FUNCTION_BLOCK SortingSafeSteps (* Standard safe-position sequence and its original timing. *)
  (* Standard: 61499-2 *)
  (* Version 3.0, 2026-11-12, sorting2n, sorting2n *)
  PACKAGE Main;
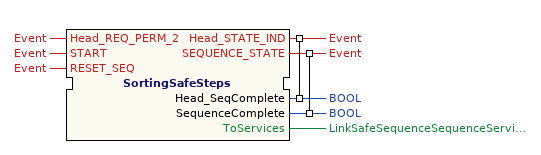
  EVENT_INPUT
    Head_REQ_PERM_2;
    START;
    RESET_SEQ;
  END_EVENT
  EVENT_OUTPUT
    Head_STATE_IND WITH Head_SeqComplete;
    SEQUENCE_STATE WITH SequenceComplete;
  END_EVENT
  VAR_OUTPUT
    Head_SeqComplete : BOOL;
    SequenceComplete : BOOL;
  END_VAR
  PLUGS
    ToServices : LinkSafeSequenceSequenceServices;
  END_PLUGS
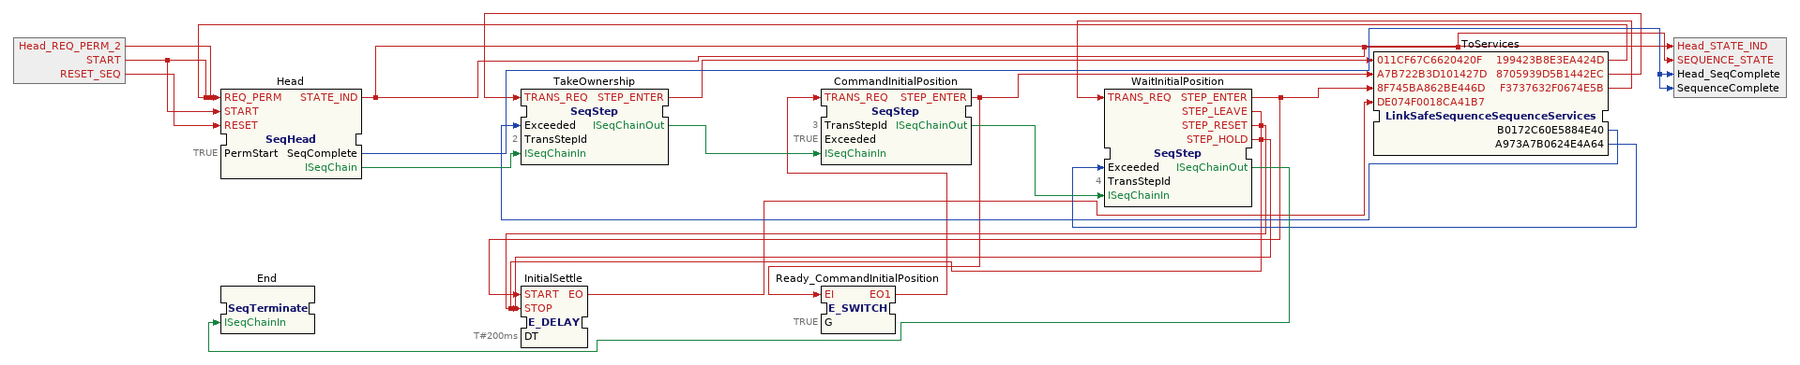
  FBS
    Head : SeqHead(PermStart := TRUE);
    End : SeqTerminate;
    TakeOwnership : SeqStep(TransStepId := 2);
    CommandInitialPosition : SeqStep(TransStepId := 3, Exceeded := TRUE);
    WaitInitialPosition : SeqStep(TransStepId := 4);
    InitialSettle : E_DELAY(DT := T#200ms);
    Ready_CommandInitialPosition : E_SWITCH(G := TRUE);
  END_FBS
  EVENT_CONNECTIONS
    Head.STATE_IND TO Head_STATE_IND;
    ToServices.199423B8E3EA424D TO Head.REQ_PERM;
    Head_REQ_PERM_2 TO Head.REQ_PERM;
    TakeOwnership.STEP_ENTER TO ToServices.011CF67C6620420F;
    ToServices.8705939D5B1442EC TO TakeOwnership.TRANS_REQ;
    CommandInitialPosition.STEP_ENTER TO ToServices.A7B722B3D101427D;
    CommandInitialPosition.STEP_ENTER TO Ready_CommandInitialPosition.EI;
    Ready_CommandInitialPosition.EO1 TO CommandInitialPosition.TRANS_REQ;
    WaitInitialPosition.STEP_ENTER TO ToServices.8F745BA862BE446D;
    WaitInitialPosition.STEP_ENTER TO InitialSettle.START;
    InitialSettle.EO TO ToServices.DE074F0018CA41B7;
    WaitInitialPosition.STEP_LEAVE TO InitialSettle.STOP;
    WaitInitialPosition.STEP_RESET TO InitialSettle.STOP;
    WaitInitialPosition.STEP_HOLD TO InitialSettle.STOP;
    ToServices.F3737632F0674E5B TO WaitInitialPosition.TRANS_REQ;
    START TO Head.REQ_PERM;
    START TO Head.START;
    RESET_SEQ TO Head.RESET;
    Head.STATE_IND TO SEQUENCE_STATE;
  END_CONNECTIONS
  DATA_CONNECTIONS
    Head.SeqComplete TO Head_SeqComplete;
    ToServices.B0172C60E5884E40 TO TakeOwnership.Exceeded;
    ToServices.A973A7B0624E4A64 TO WaitInitialPosition.Exceeded;
    Head.SeqComplete TO SequenceComplete;
  END_CONNECTIONS
  ADAPTER_CONNECTIONS
    Head.ISeqChain TO TakeOwnership.ISeqChainIn;
    TakeOwnership.ISeqChainOut TO CommandInitialPosition.ISeqChainIn;
    CommandInitialPosition.ISeqChainOut TO WaitInitialPosition.ISeqChainIn;
    WaitInitialPosition.ISeqChainOut TO End.ISeqChainIn;
  END_CONNECTIONS
END_FUNCTION_BLOCK
